TYPE ST_STOEBERSI6SC6CIA402_REF_1 : FB_STOEBERSI6SC6CIA402_REF;
END_TYPE

(* stored: Version 1.1.0.1, ProductVersion 3.1.4024.15
   DUT ST_STOEBERSI6SC6CIA402_REF_1: Id {37fed269-f954-45cd-96cd-5d7f1c408a66} *)
